(* IEC 61131-3 sources: llm-plc-st-eval/data/processed_definitivo/gemini-3.1-pro-preview/B5/few_shot, 3 files *)

(* ---- ejec_1.st ---- *)
FUNCTION_BLOCK FB_Ventilador
VAR_INPUT
    quemadorOn : BOOL; (* Estado del quemador *)
END_VAR
VAR_OUTPUT
    ventilador : BOOL; (* Ventilador de enfriamiento *)
END_VAR
VAR
    tRetardoApagado : TOF; (* Temporizador de retardo a la desconexion *)
END_VAR

(* El ventilador continua funcionando 30 s despues de que se apaga el quemador *)
tRetardoApagado(IN := quemadorOn, PT := T#30S);
ventilador := tRetardoApagado.Q;
END_FUNCTION_BLOCK

(* ---- ejec_2.st ---- *)
FUNCTION_BLOCK FB_Ventilador
VAR_INPUT
    quemadorOn : BOOL; (* Estado del quemador *)
END_VAR
VAR_OUTPUT
    ventilador : BOOL; (* Ventilador de enfriamiento *)
END_VAR
VAR
    tRetardoApagado : TOF; (* Temporizador de retardo a la desconexion *)
END_VAR

(* El ventilador se mantiene encendido 30 s despues de apagarse el quemador *)
tRetardoApagado(IN := quemadorOn, PT := T#30S);
ventilador := tRetardoApagado.Q;
END_FUNCTION_BLOCK

(* ---- ejec_3.st ---- *)
FUNCTION_BLOCK FB_Ventilador
VAR_INPUT
    quemadorOn : BOOL; (* Estado del quemador *)
END_VAR
VAR_OUTPUT
    ventilador : BOOL; (* Ventilador de enfriamiento *)
END_VAR
VAR
    tRetardoApagado : TOF; (* Temporizador de retardo a la desconexion *)
END_VAR

(* El ventilador continua encendido 30 s despues de apagarse el quemador *)
tRetardoApagado(IN := quemadorOn, PT := T#30S);
ventilador := tRetardoApagado.Q;
END_FUNCTION_BLOCK
